// TIA Portal V14 SP1 export
// export: Created 2000-01-01T00:00:00.0000000Z, ExportSetting None
DATA_BLOCK "MCP_RC_DB7"   // DB9807
{ S7_Optimized_Access := 'TRUE' }
   VAR
      Aa : Int := 1;
      R : Real := 1.5;
      W : Int := 3;
      Motor : "MCP_RC_UDT";
   END_VAR
BEGIN
END_DATA_BLOCK
